Fanuc KAREL source: KB00109.KL

PROGRAM KB00109
%NOLOCKGROUP
VAR
  P1: POSITION
  RESULT: POSITION
BEGIN
  RESULT = INV(P1)
END KB00109
